(* Logix 5000 project; controller NWGG 1756-L72 rev 35.12; software revision 35.00; part 5 of 19 *)
(* tags used below, declared in another part *)
   _101AUTO : ALIAS FOR B9[101].4;
   _101HAND : ALIAS FOR B9[101].3;
   _101M : ALIAS FOR O25[9].3;
   _101MB : ALIAS FOR B9[101].2;
   _101STB : ALIAS FOR B9[101].0;
   _101STPB : ALIAS FOR B9[101].1;
   _101Y : ALIAS FOR I25[1].3;
   _102AUTO : ALIAS FOR B9[102].4;
   _102HAND : ALIAS FOR B9[102].3;
   _102M : ALIAS FOR O25[8].9;
   _102MB : ALIAS FOR B9[102].2;
   _102STB : ALIAS FOR B9[102].0;
   _102STPB : ALIAS FOR B9[102].1;
   _102Y : ALIAS FOR I25[0].9;
   _103AUTO : ALIAS FOR B9[103].4;
   _103HAND : ALIAS FOR B9[103].3;
   _103M : ALIAS FOR O25[8].12;
   _103MB : ALIAS FOR B9[103].2;
   _103STB : ALIAS FOR B9[103].0;
   _103STPB : ALIAS FOR B9[103].1;
   _103Y : ALIAS FOR I25[0].12;
   _106AUTO : ALIAS FOR B9[106].4;
   _106HAND : ALIAS FOR B9[106].3;
   _106M : ALIAS FOR O25[9].5;
   _106MB : ALIAS FOR B9[106].2;
   _106Y : ALIAS FOR I25[1].5;
   _107AUTO : ALIAS FOR B9[107].4;
   _107HAND : ALIAS FOR B9[107].3;
   _107M : ALIAS FOR O25[9].12;
   _107MB : ALIAS FOR B9[107].2;
   _107PS : ALIAS FOR I25[4].2;
   _107PSB : ALIAS FOR B9[107].5;
   _107STB : ALIAS FOR B9[107].0;
   _107STPB : ALIAS FOR B9[107].1;
   _107Y : ALIAS FOR I25[1].12;
   _108AUTO : ALIAS FOR B9[108].4;
   _108HAND : ALIAS FOR B9[108].3;
   _108M : ALIAS FOR O25[10].15;
   _108MB : ALIAS FOR B9[108].2;
   _108PS : ALIAS FOR I25[4].1;
   _108STB : ALIAS FOR B9[108].0;
   _108STPB : ALIAS FOR B9[108].1;
   _108Y : ALIAS FOR I25[2].15;
   _109_PS_DLY : ALIAS FOR T11[4];
   _109_SLOW_D : ALIAS FOR T11[5];
   _109_SLW_SP : ALIAS FOR I25[3].14;
   _109_STOP_D : ALIAS FOR T11[6];
   _109_STP_SP : ALIAS FOR I25[3].15;
   _109AUTO : ALIAS FOR B9[109].4;
   _109HAND : ALIAS FOR B9[109].3;
   _109M : ALIAS FOR O25[10].9;
   _109MB : ALIAS FOR B9[109].2;
   _109PS : ALIAS FOR I25[4].0;
   _109STB : ALIAS FOR B9[109].0;
   _109STPB : ALIAS FOR B9[109].1;
   _109Y : ALIAS FOR I25[2].9;
   _110AUTO : ALIAS FOR B9[110].4;
   _110HAND : ALIAS FOR B9[110].3;
   _110M : ALIAS FOR O25[8].15;
   _110MB : ALIAS FOR B9[110].2;
   _110STB : ALIAS FOR B9[110].0;
   _110STPB : ALIAS FOR B9[110].1;
   _110Y : ALIAS FOR I25[0].15;
   _111AUTO : ALIAS FOR B9[111].4;
   _111HAND : ALIAS FOR B9[111].3;
   _111M : ALIAS FOR O25[9].0;
   _111MB : ALIAS FOR B9[111].2;
   _111STB : ALIAS FOR B9[111].0;
   _111STPB : ALIAS FOR B9[111].1;
   _111Y : ALIAS FOR I25[1].0;
   _113AUTO : ALIAS FOR B9[113].4;
   _113HAND : ALIAS FOR B9[113].3;
   _113M : ALIAS FOR O25[10].5;
   _113MB : ALIAS FOR B9[113].2;
   _113STB : ALIAS FOR B9[113].0;
   _113STPB : ALIAS FOR B9[113].1;
   _113Y : ALIAS FOR I25[2].5;
   _116AUTO : ALIAS FOR B9[116].4;
   _116HAND : ALIAS FOR B9[116].3;
   _116M : ALIAS FOR O25[10].10;
   _116MB : ALIAS FOR B9[116].2;
   _116STB : ALIAS FOR B9[116].0;
   _116STPB : ALIAS FOR B9[116].1;
   _116Y : ALIAS FOR I25[2].10;
   _117AUTO : ALIAS FOR B9[117].4;
   _117HAND : ALIAS FOR B9[117].3;
   _117M : ALIAS FOR O25[10].8;
   _117MB : ALIAS FOR B9[117].2;
   _117STB : ALIAS FOR B9[117].0;
   _117STPB : ALIAS FOR B9[117].1;
   _117Y : ALIAS FOR I25[2].8;
   _11_PS : ALIAS FOR I25[4].14;
   _11_PS_DLY : ALIAS FOR T11[2];
   _11_SLOW_SP : ALIAS FOR I25[4].3;
   _11_STOP_SP : ALIAS FOR I25[4].6;
   _11AUTO : ALIAS FOR B9[11].4;
   _11HAND : ALIAS FOR B9[11].3;
   _11M : ALIAS FOR O25[9].2;
   _11MB : ALIAS FOR B9[11].2;
   _11STB : ALIAS FOR B9[11].0;
   _11STPB : ALIAS FOR B9[11].1;
   _11Y : ALIAS FOR I25[1].2;
   _122AUTO : ALIAS FOR B9[122].4;
   _122HAND : ALIAS FOR B9[122].3;
   _122M : ALIAS FOR O25[9].1;
   _122MB : ALIAS FOR B9[122].2;
   _122STB : ALIAS FOR B9[122].0;
   _122STPB : ALIAS FOR B9[122].1;
   _122Y : ALIAS FOR I25[1].1;
   _123_COMPUW : ALIAS FOR I18[7];
   _123_COMPUW1 : ALIAS FOR N7[20];
   _123AUTO : ALIAS FOR B9[123].4;
   _123HAND : ALIAS FOR B9[123].3;
   _123M : ALIAS FOR O25[10].6;
   _123MB : ALIAS FOR B9[123].2;
   _123STB : ALIAS FOR B9[123].0;
   _123STPB : ALIAS FOR B9[123].1;
   _123Y : ALIAS FOR I25[2].6;
   _124M : ALIAS FOR O25[9].13;
   _1AUTO : ALIAS FOR B9[1].4;
   _1HAND : ALIAS FOR B9[1].3;
   _1M : ALIAS FOR O25[9].8;
   _1MB : ALIAS FOR B9[1].2;
   _1STB : ALIAS FOR B9[1].0;
   _1STPB : ALIAS FOR B9[1].1;
   _1Y : ALIAS FOR I25[1].8;
   _25_16_0 : ALIAS FOR N200[10];
   _25_16_1 : ALIAS FOR N200[11];
   _25_16_2 : ALIAS FOR N200[12];
   _25_16_3 : ALIAS FOR N200[13];
   _2AUTO : ALIAS FOR B9[2].4;
   _2HAND : ALIAS FOR B9[2].3;
   _2M : ALIAS FOR O25[9].15;
   _2MB : ALIAS FOR B9[2].2;
   _2STB : ALIAS FOR B9[2].0;
   _2STPB : ALIAS FOR B9[2].1;
   _2Y : ALIAS FOR I25[1].15;
   _35AUTO : ALIAS FOR B9[35].4;
   _35HAND : ALIAS FOR B9[35].3;
   _35M : ALIAS FOR O25[10].13;
   _35MB : ALIAS FOR B9[35].2;
   _35STB : ALIAS FOR B9[35].0;
   _35STPB : ALIAS FOR B9[35].1;
   _35Y : ALIAS FOR I25[2].13;
   _36_FREQ_IN : ALIAS FOR N7[1];
   _36_FREQ_OU : ALIAS FOR N7[3];
   _36_SET_SPD : ALIAS FOR N7[2];
   _36_VFD_TO : ALIAS FOR N180[0];
   _36M : ALIAS FOR O25[8].0;
   _36RAUTO : ALIAS FOR B9[36].4;
   _36RHAND : ALIAS FOR B9[36].3;
   _36RMB : ALIAS FOR B9[36].2;
   _36RSTB : ALIAS FOR B9[36].0;
   _36RSTPB : ALIAS FOR B9[36].1;
   _36Y : ALIAS FOR I25[0].0;
   _3AUTO : ALIAS FOR B9[3].4;
   _3HAND : ALIAS FOR B9[3].3;
   _3M : ALIAS FOR O25[10].0;
   _3MB : ALIAS FOR B9[3].2;
   _3STB : ALIAS FOR B9[3].0;
   _3STPB : ALIAS FOR B9[3].1;
   _3Y : ALIAS FOR I25[2].0;
   _42AUTO : ALIAS FOR B9[42].4;
   _42HAND : ALIAS FOR B9[42].3;
   _42M : ALIAS FOR O25[11].1;
   _42MB : ALIAS FOR B9[42].2;
   _42STB : ALIAS FOR B9[42].0;
   _42STPB : ALIAS FOR B9[42].1;
   _42Y : ALIAS FOR I25[3].1;
   _43_ACC_WEI : ALIAS FOR C5[1].ACC;
   _43_BINDICA : ALIAS FOR B9[43].5;
   _43_RESET_C : ALIAS FOR B9[43].6;
   _43_SCREEN : ALIAS FOR C5[1];
   _43_SCREENI : ALIAS FOR I7.14;
   _43_WEIGHT : ALIAS FOR N7[0];
   _43AUTO : ALIAS FOR B9[43].4;
   _43HAND : ALIAS FOR B9[43].3;
   _43M : ALIAS FOR O25[10].14;
   _43MB : ALIAS FOR B9[43].2;
   _43STB : ALIAS FOR B9[43].0;
   _43STPB : ALIAS FOR B9[43].1;
   _43Y : ALIAS FOR I25[2].14;
   _47AUTO : ALIAS FOR B9[47].4;
   _47HAND : ALIAS FOR B9[47].3;
   _47M : ALIAS FOR O25[9].10;
   _47MB : ALIAS FOR B9[47].2;
   _47STB : ALIAS FOR B9[47].0;
   _47STPB : ALIAS FOR B9[47].1;
   _47Y : ALIAS FOR I25[1].10;
   _48_FREQ_IN : ALIAS FOR N7[10];
   _48_FREQ_OU : ALIAS FOR N7[12];
   _48_SET_SPD : ALIAS FOR N7[11];
   _48_VFD_TO : ALIAS FOR N180[2];
   _48AUTO : ALIAS FOR B9[48].4;
   _48HAND : ALIAS FOR B9[48].3;
   _48M : ALIAS FOR O25[8].3;
   _48MB : ALIAS FOR B9[48].2;
   _48STB : ALIAS FOR B9[48].0;
   _48STPB : ALIAS FOR B9[48].1;
   _48Y : ALIAS FOR I25[0].3;
   _49AUTO : ALIAS FOR B9[49].4;
   _49HAND : ALIAS FOR B9[49].3;
   _49M : ALIAS FOR O25[9].9;
   _49MB : ALIAS FOR B9[49].2;
   _49STB : ALIAS FOR B9[49].0;
   _49STPB : ALIAS FOR B9[49].1;
   _49Y : ALIAS FOR I25[1].9;
   _4AUTO : ALIAS FOR B9[4].4;
   _4HAND : ALIAS FOR B9[4].3;
   _4M : ALIAS FOR O25[10].1;
   _4MB : ALIAS FOR B9[4].2;
   _4STB : ALIAS FOR B9[4].0;
   _4STPB : ALIAS FOR B9[4].1;
   _4Y : ALIAS FOR I25[2].1;
   _50AUTO : ALIAS FOR B9[50].4;
   _50HAND : ALIAS FOR B9[50].3;
   _50M : ALIAS FOR O25[8].14;
   _50MB : ALIAS FOR B9[50].2;
   _50STB : ALIAS FOR B9[50].0;
   _50STPB : ALIAS FOR B9[50].1;
   _50Y : ALIAS FOR I25[0].14;
   _51_FREQ_IN : ALIAS FOR N7[13];
   _51_FREQ_OU : ALIAS FOR N7[15];
   _51_SET_SPD : ALIAS FOR N7[14];
   _51_VFD_TO : ALIAS FOR N180[3];
   _51AUTO : ALIAS FOR B9[51].4;
   _51HAND : ALIAS FOR B9[51].3;
   _51M : ALIAS FOR O25[8].4;
   _51MB : ALIAS FOR B9[51].2;
   _51STB : ALIAS FOR B9[51].0;
   _51STPB : ALIAS FOR B9[51].1;
   _51Y : ALIAS FOR I25[0].4;
   _52_FREQ_IN : ALIAS FOR N7[16];
   _52_FREQ_OU : ALIAS FOR N7[18];
   _52_SET_SPD : ALIAS FOR N7[17];
   _52AUTO : ALIAS FOR B9[52].4;
   _52HAND : ALIAS FOR B9[52].3;
   _52M : ALIAS FOR O25[8].6;
   _52MB : ALIAS FOR B9[52].2;
   _52STB : ALIAS FOR B9[52].0;
   _52STPB : ALIAS FOR B9[52].1;
   _52Y : ALIAS FOR I25[0].6;
   _53_FREQ_IN : ALIAS FOR N7[7];
   _53_FREQ_OU : ALIAS FOR N7[9];
   _53_SET_SPD : ALIAS FOR N7[8];
   _53_VFD_TO : ALIAS FOR N180[1];
   _53AUTO : ALIAS FOR B9[53].4;
   _53HAND : ALIAS FOR B9[53].3;
   _53M : ALIAS FOR O25[8].2;
   _53MB : ALIAS FOR B9[53].2;
(* _2_MAIN, continued *)

ROUTINE _09_SEED_MTR_9   (* ladder *)
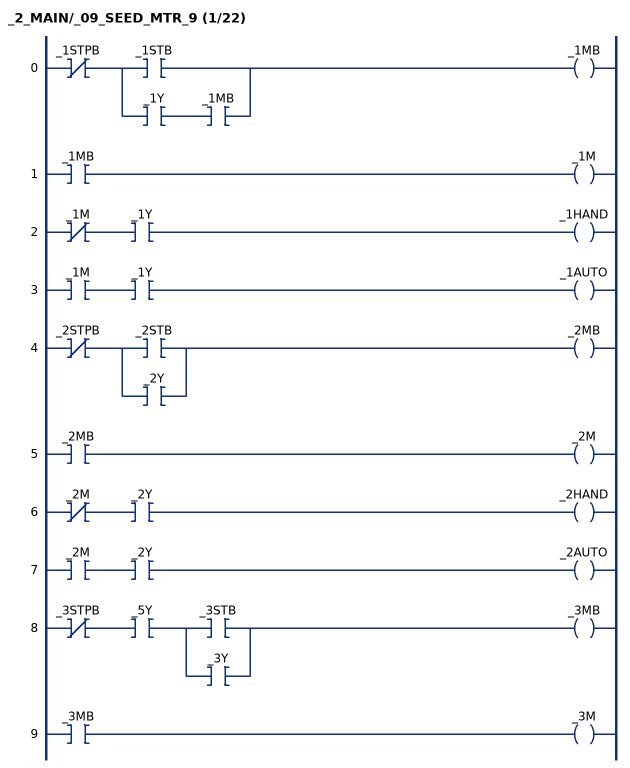
   0: XIO(_1STPB)[XIC(_1STB) ,XIC(_1Y) XIC(_1MB) ]OTE(_1MB);
   1: XIC(_1MB)OTE(_1M);
   2: XIO(_1M)XIC(_1Y)OTE(_1HAND);
   3: XIC(_1M)XIC(_1Y)OTE(_1AUTO);
   4: XIO(_2STPB)[XIC(_2STB) ,XIC(_2Y) ]OTE(_2MB);
   5: XIC(_2MB)OTE(_2M);
   6: XIO(_2M)XIC(_2Y)OTE(_2HAND);
   7: XIC(_2M)XIC(_2Y)OTE(_2AUTO);
   8: XIO(_3STPB)XIC(_5Y)[XIC(_3STB) ,XIC(_3Y) ]OTE(_3MB);
   9: XIC(_3MB)OTE(_3M);
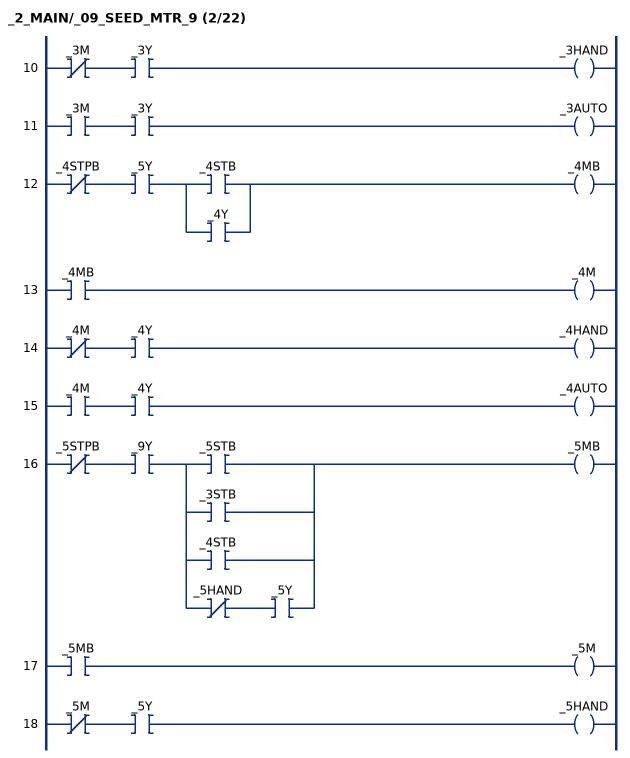
   10: XIO(_3M)XIC(_3Y)OTE(_3HAND);
   11: XIC(_3M)XIC(_3Y)OTE(_3AUTO);
   12: XIO(_4STPB)XIC(_5Y)[XIC(_4STB) ,XIC(_4Y) ]OTE(_4MB);
   13: XIC(_4MB)OTE(_4M);
   14: XIO(_4M)XIC(_4Y)OTE(_4HAND);
   15: XIC(_4M)XIC(_4Y)OTE(_4AUTO);
   16: XIO(_5STPB)XIC(_9Y)[XIC(_5STB) ,XIC(_3STB) ,XIC(_4STB) ,XIO(_5HAND) XIC(_5Y) ]OTE(_5MB);
   17: XIC(_5MB)OTE(_5M);
   18: XIO(_5M)XIC(_5Y)OTE(_5HAND);
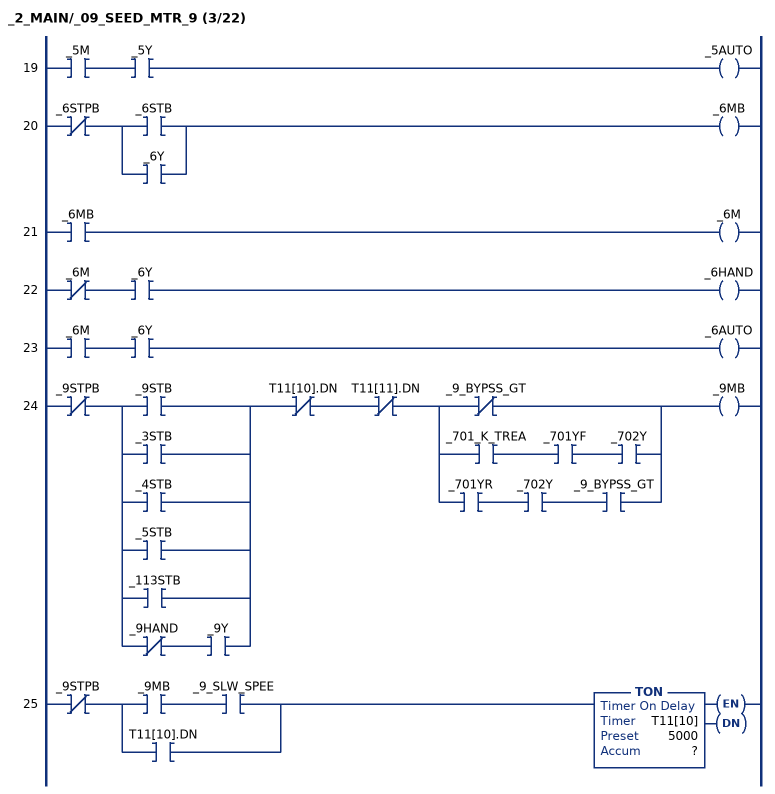
   19: XIC(_5M)XIC(_5Y)OTE(_5AUTO);
   20: XIO(_6STPB)[XIC(_6STB) ,XIC(_6Y) ]OTE(_6MB);
   21: XIC(_6MB)OTE(_6M);
   22: XIO(_6M)XIC(_6Y)OTE(_6HAND);
   23: XIC(_6M)XIC(_6Y)OTE(_6AUTO);
   24: XIO(_9STPB)[XIC(_9STB) ,XIC(_3STB) ,XIC(_4STB) ,XIC(_5STB) ,XIC(_113STB) ,XIO(_9HAND) XIC(_9Y) ]XIO(T11[10].DN)XIO(T11[11].DN)[XIO(_9_BYPSS_GT) ,XIC(_701_K_TREA) XIC(_701YF) XIC(_702Y) ,XIC(_701YR) XIC(_702Y) XIC(_9_BYPSS_GT) ]OTE(_9MB);
   25: XIO(_9STPB)[XIC(_9MB) XIC(_9_SLW_SPEE) ,XIC(T11[10].DN) ]TON(T11[10],?,?);
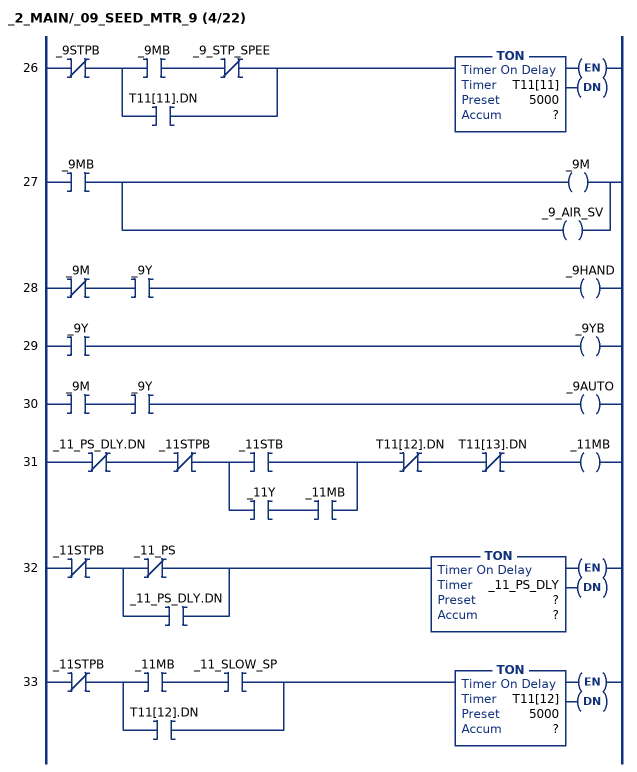
   26: XIO(_9STPB)[XIC(_9MB) XIO(_9_STP_SPEE) ,XIC(T11[11].DN) ]TON(T11[11],?,?);
   27: XIC(_9MB)[OTE(_9M) ,OTE(_9_AIR_SV) ];
   28: XIO(_9M)XIC(_9Y)OTE(_9HAND);
   29: XIC(_9Y)OTE(_9YB);
   30: XIC(_9M)XIC(_9Y)OTE(_9AUTO);
   31: XIO(_11_PS_DLY.DN)XIO(_11STPB)[XIC(_11STB) ,XIC(_11Y) XIC(_11MB) ]XIO(T11[12].DN)XIO(T11[13].DN)OTE(_11MB);
   32: XIO(_11STPB)[XIO(_11_PS) ,XIC(_11_PS_DLY.DN) ]TON(_11_PS_DLY,?,?);
   33: XIO(_11STPB)[XIC(_11MB) XIC(_11_SLOW_SP) ,XIC(T11[12].DN) ]TON(T11[12],?,?);
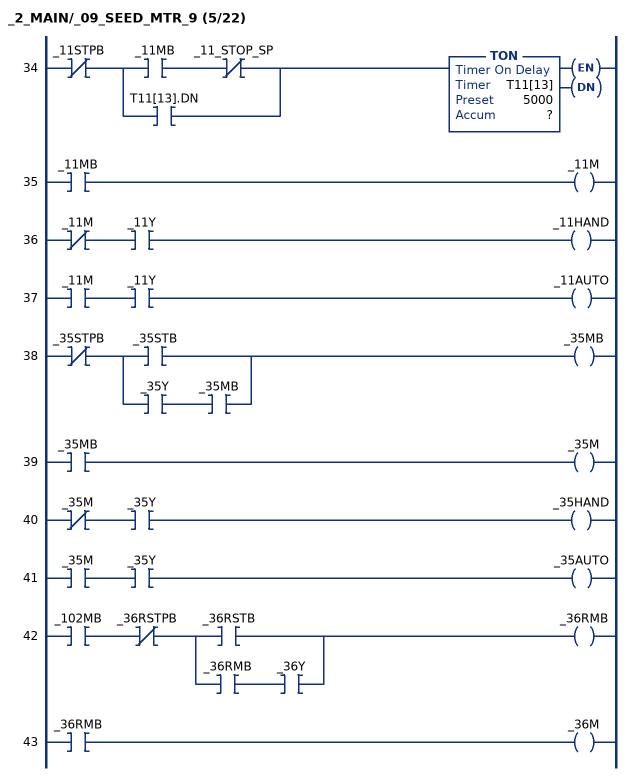
   34: XIO(_11STPB)[XIC(_11MB) XIO(_11_STOP_SP) ,XIC(T11[13].DN) ]TON(T11[13],?,?);
   35: XIC(_11MB)OTE(_11M);
   36: XIO(_11M)XIC(_11Y)OTE(_11HAND);
   37: XIC(_11M)XIC(_11Y)OTE(_11AUTO);
   38: XIO(_35STPB)[XIC(_35STB) ,XIC(_35Y) XIC(_35MB) ]OTE(_35MB);
   39: XIC(_35MB)OTE(_35M);
   40: XIO(_35M)XIC(_35Y)OTE(_35HAND);
   41: XIC(_35M)XIC(_35Y)OTE(_35AUTO);
   42: XIC(_102MB)XIO(_36RSTPB)[XIC(_36RSTB) ,XIC(_36RMB) XIC(_36Y) ]OTE(_36RMB);
   43: XIC(_36RMB)OTE(_36M);
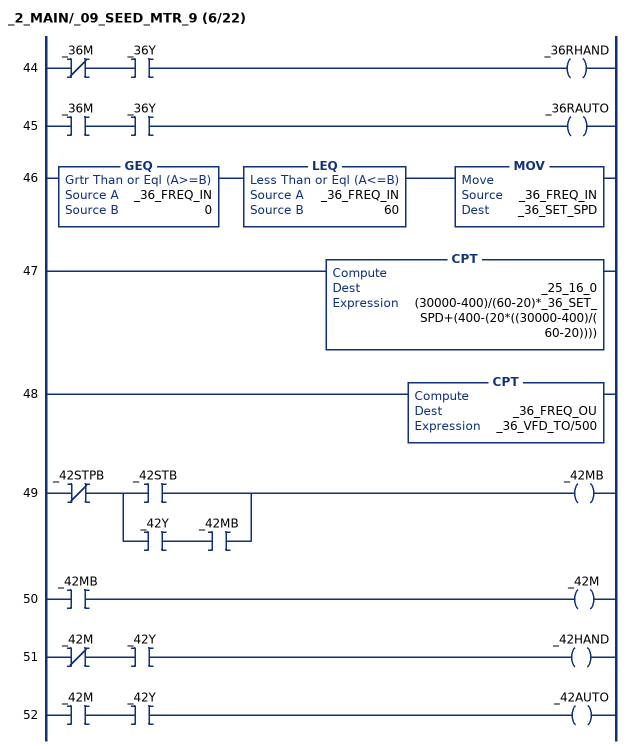
   44: XIO(_36M)XIC(_36Y)OTE(_36RHAND);
   45: XIC(_36M)XIC(_36Y)OTE(_36RAUTO);
   46: GEQ(_36_FREQ_IN,0)LEQ(_36_FREQ_IN,60)MOV(_36_FREQ_IN,_36_SET_SPD);
   47: CPT(_25_16_0,(30000-400)/(60-20)*_36_SET_SPD+(400-(20*((30000-400)/(60-20)))));
   48: CPT(_36_FREQ_OU,_36_VFD_TO/500);
   49: XIO(_42STPB)[XIC(_42STB) ,XIC(_42Y) XIC(_42MB) ]OTE(_42MB);
   50: XIC(_42MB)OTE(_42M);
   51: XIO(_42M)XIC(_42Y)OTE(_42HAND);
   52: XIC(_42M)XIC(_42Y)OTE(_42AUTO);
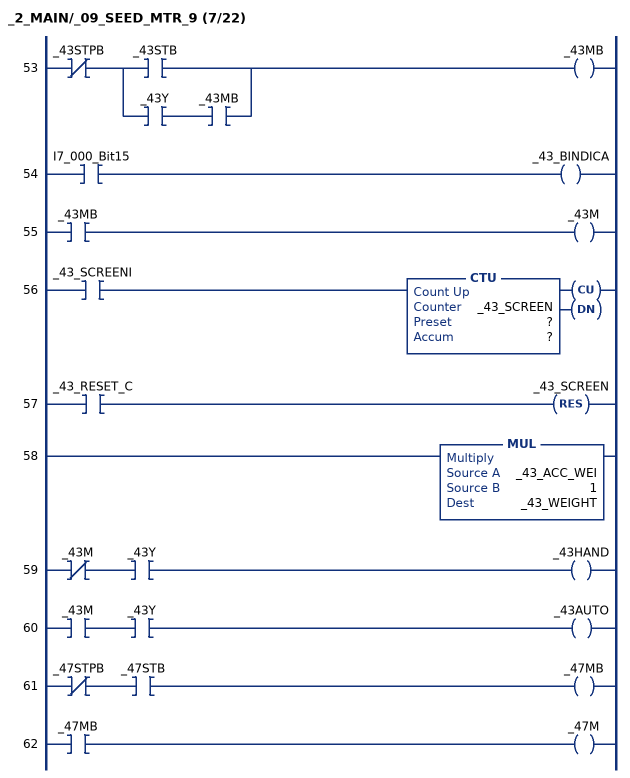
   53: XIO(_43STPB)[XIC(_43STB) ,XIC(_43Y) XIC(_43MB) ]OTE(_43MB);
   54: XIC(I7_000_Bit15)OTE(_43_BINDICA);
   55: XIC(_43MB)OTE(_43M);
   56: XIC(_43_SCREENI)CTU(_43_SCREEN,?,?);
   57: XIC(_43_RESET_C)RES(_43_SCREEN);
   58: MUL(_43_ACC_WEI,1,_43_WEIGHT);
   59: XIO(_43M)XIC(_43Y)OTE(_43HAND);
   60: XIC(_43M)XIC(_43Y)OTE(_43AUTO);
   61: XIO(_47STPB)XIC(_47STB)OTE(_47MB);
   62: XIC(_47MB)OTE(_47M);
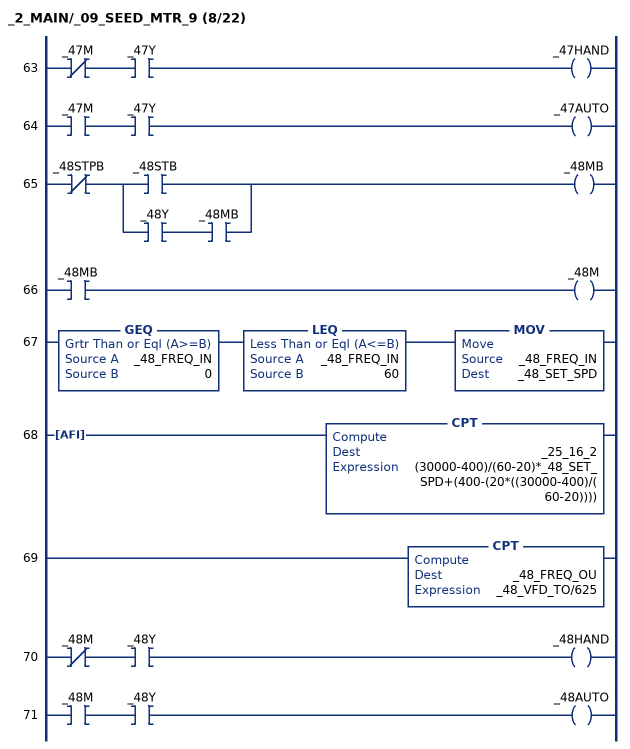
   63: XIO(_47M)XIC(_47Y)OTE(_47HAND);
   64: XIC(_47M)XIC(_47Y)OTE(_47AUTO);
   65: XIO(_48STPB)[XIC(_48STB) ,XIC(_48Y) XIC(_48MB) ]OTE(_48MB);
   66: XIC(_48MB)OTE(_48M);
   67: GEQ(_48_FREQ_IN,0)LEQ(_48_FREQ_IN,60)MOV(_48_FREQ_IN,_48_SET_SPD);
   68: AFI()CPT(_25_16_2,(30000-400)/(60-20)*_48_SET_SPD+(400-(20*((30000-400)/(60-20)))));
   69: CPT(_48_FREQ_OU,_48_VFD_TO/625);
   70: XIO(_48M)XIC(_48Y)OTE(_48HAND);
   71: XIC(_48M)XIC(_48Y)OTE(_48AUTO);
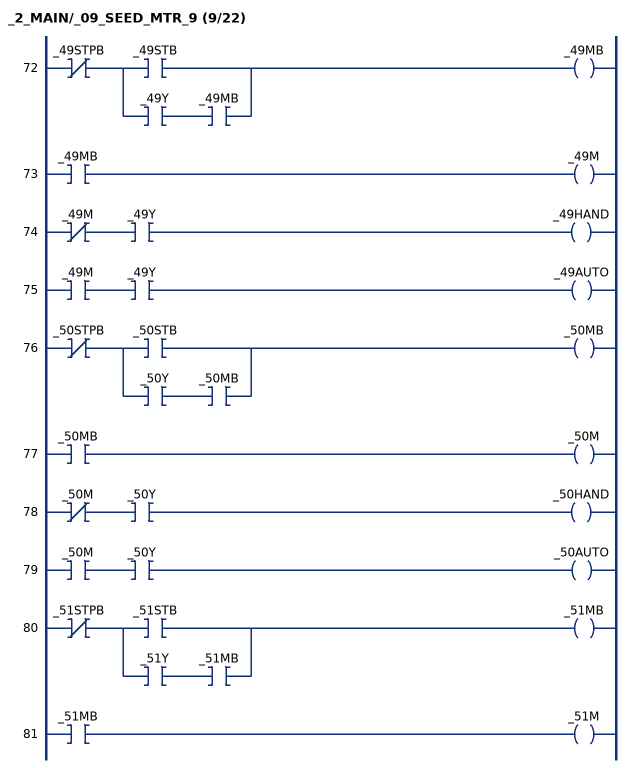
   72: XIO(_49STPB)[XIC(_49STB) ,XIC(_49Y) XIC(_49MB) ]OTE(_49MB);
   73: XIC(_49MB)OTE(_49M);
   74: XIO(_49M)XIC(_49Y)OTE(_49HAND);
   75: XIC(_49M)XIC(_49Y)OTE(_49AUTO);
   76: XIO(_50STPB)[XIC(_50STB) ,XIC(_50Y) XIC(_50MB) ]OTE(_50MB);
   77: XIC(_50MB)OTE(_50M);
   78: XIO(_50M)XIC(_50Y)OTE(_50HAND);
   79: XIC(_50M)XIC(_50Y)OTE(_50AUTO);
   80: XIO(_51STPB)[XIC(_51STB) ,XIC(_51Y) XIC(_51MB) ]OTE(_51MB);
   81: XIC(_51MB)OTE(_51M);
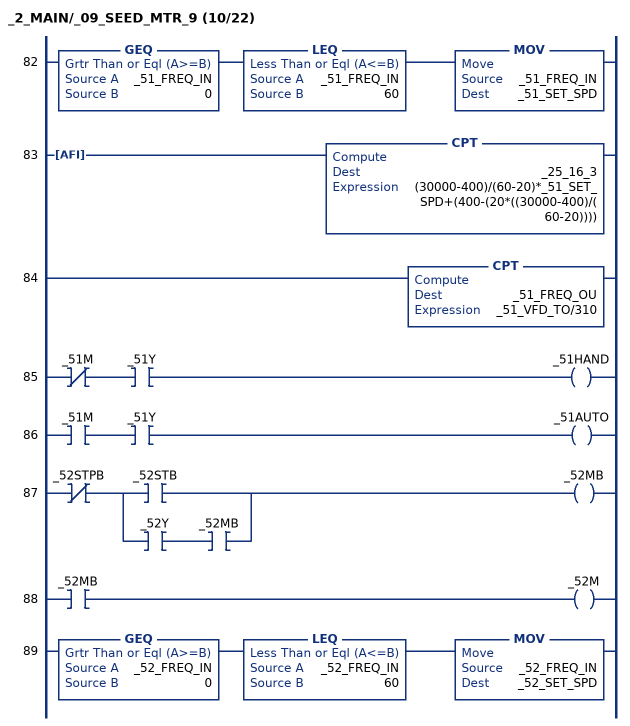
   82: GEQ(_51_FREQ_IN,0)LEQ(_51_FREQ_IN,60)MOV(_51_FREQ_IN,_51_SET_SPD);
   83: AFI()CPT(_25_16_3,(30000-400)/(60-20)*_51_SET_SPD+(400-(20*((30000-400)/(60-20)))));
   84: CPT(_51_FREQ_OU,_51_VFD_TO/310);
   85: XIO(_51M)XIC(_51Y)OTE(_51HAND);
   86: XIC(_51M)XIC(_51Y)OTE(_51AUTO);
   87: XIO(_52STPB)[XIC(_52STB) ,XIC(_52Y) XIC(_52MB) ]OTE(_52MB);
   88: XIC(_52MB)OTE(_52M);
   89: GEQ(_52_FREQ_IN,0)LEQ(_52_FREQ_IN,60)MOV(_52_FREQ_IN,_52_SET_SPD);
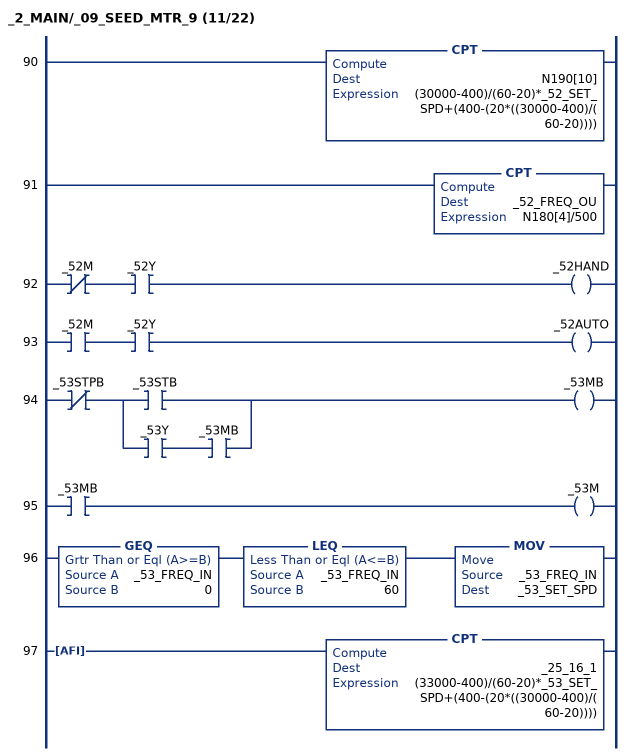
   90: CPT(N190[10],(30000-400)/(60-20)*_52_SET_SPD+(400-(20*((30000-400)/(60-20)))));
   91: CPT(_52_FREQ_OU,N180[4]/500);
   92: XIO(_52M)XIC(_52Y)OTE(_52HAND);
   93: XIC(_52M)XIC(_52Y)OTE(_52AUTO);
   94: XIO(_53STPB)[XIC(_53STB) ,XIC(_53Y) XIC(_53MB) ]OTE(_53MB);
   95: XIC(_53MB)OTE(_53M);
   96: GEQ(_53_FREQ_IN,0)LEQ(_53_FREQ_IN,60)MOV(_53_FREQ_IN,_53_SET_SPD);
   97: AFI()CPT(_25_16_1,(33000-400)/(60-20)*_53_SET_SPD+(400-(20*((30000-400)/(60-20)))));
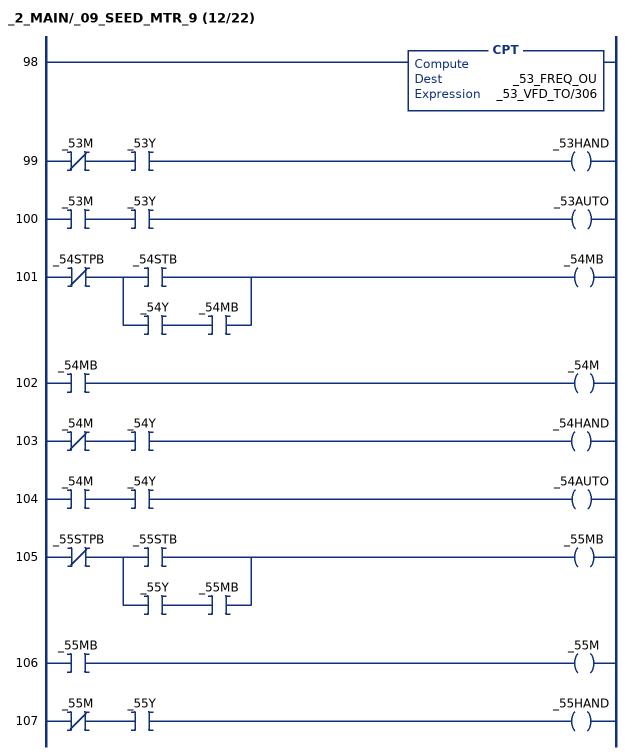
   98: CPT(_53_FREQ_OU,_53_VFD_TO/306);
   99: XIO(_53M)XIC(_53Y)OTE(_53HAND);
   100: XIC(_53M)XIC(_53Y)OTE(_53AUTO);
   101: XIO(_54STPB)[XIC(_54STB) ,XIC(_54Y) XIC(_54MB) ]OTE(_54MB);
   102: XIC(_54MB)OTE(_54M);
   103: XIO(_54M)XIC(_54Y)OTE(_54HAND);
   104: XIC(_54M)XIC(_54Y)OTE(_54AUTO);
   105: XIO(_55STPB)[XIC(_55STB) ,XIC(_55Y) XIC(_55MB) ]OTE(_55MB);
   106: XIC(_55MB)OTE(_55M);
   107: XIO(_55M)XIC(_55Y)OTE(_55HAND);
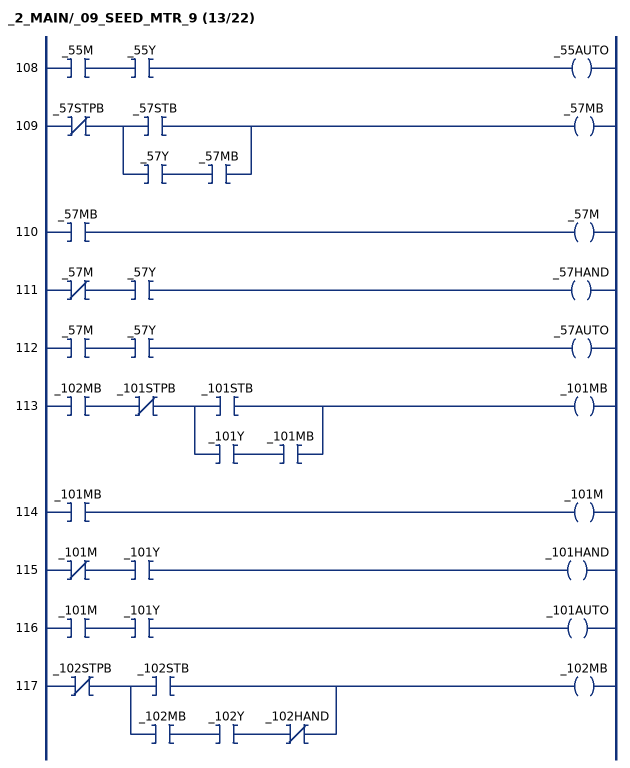
   108: XIC(_55M)XIC(_55Y)OTE(_55AUTO);
   109: XIO(_57STPB)[XIC(_57STB) ,XIC(_57Y) XIC(_57MB) ]OTE(_57MB);
   110: XIC(_57MB)OTE(_57M);
   111: XIO(_57M)XIC(_57Y)OTE(_57HAND);
   112: XIC(_57M)XIC(_57Y)OTE(_57AUTO);
   113: XIC(_102MB)XIO(_101STPB)[XIC(_101STB) ,XIC(_101Y) XIC(_101MB) ]OTE(_101MB);
   114: XIC(_101MB)OTE(_101M);
   115: XIO(_101M)XIC(_101Y)OTE(_101HAND);
   116: XIC(_101M)XIC(_101Y)OTE(_101AUTO);
   117: XIO(_102STPB)[XIC(_102STB) ,XIC(_102MB) XIC(_102Y) XIO(_102HAND) ]OTE(_102MB);
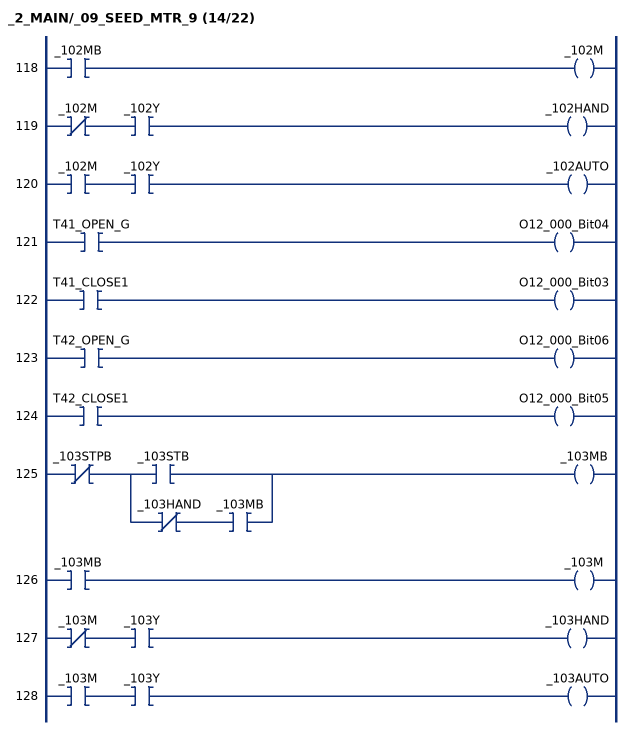
   118: XIC(_102MB)OTE(_102M);
   119: XIO(_102M)XIC(_102Y)OTE(_102HAND);
   120: XIC(_102M)XIC(_102Y)OTE(_102AUTO);
   121: XIC(T41_OPEN_G)OTE(O12_000_Bit04);
   122: XIC(T41_CLOSE1)OTE(O12_000_Bit03);
   123: XIC(T42_OPEN_G)OTE(O12_000_Bit06);
   124: XIC(T42_CLOSE1)OTE(O12_000_Bit05);
   125: XIO(_103STPB)[XIC(_103STB) ,XIO(_103HAND) XIC(_103MB) ]OTE(_103MB);
   126: XIC(_103MB)OTE(_103M);
   127: XIO(_103M)XIC(_103Y)OTE(_103HAND);
   128: XIC(_103M)XIC(_103Y)OTE(_103AUTO);
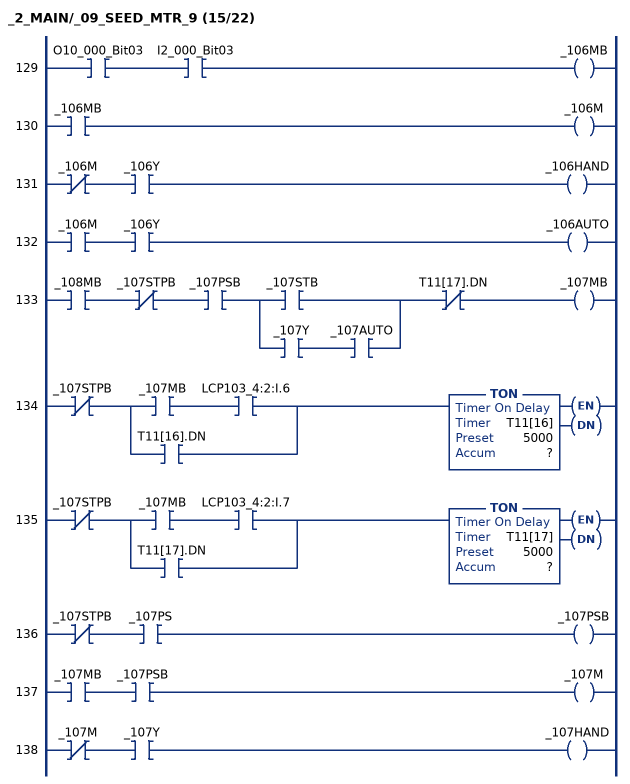
   129: XIC(O10_000_Bit03)XIC(I2_000_Bit03)OTE(_106MB);
   130: XIC(_106MB)OTE(_106M);
   131: XIO(_106M)XIC(_106Y)OTE(_106HAND);
   132: XIC(_106M)XIC(_106Y)OTE(_106AUTO);
   133: XIC(_108MB)XIO(_107STPB)XIC(_107PSB)[XIC(_107STB) ,XIC(_107Y) XIC(_107AUTO) ]XIO(T11[17].DN)OTE(_107MB);
   134: XIO(_107STPB)[XIC(_107MB) XIC(LCP103_4:2:I.6) ,XIC(T11[16].DN) ]TON(T11[16],?,?);
   135: XIO(_107STPB)[XIC(_107MB) XIC(LCP103_4:2:I.7) ,XIC(T11[17].DN) ]TON(T11[17],?,?);
   136: XIO(_107STPB)XIC(_107PS)OTE(_107PSB);
   137: XIC(_107MB)XIC(_107PSB)OTE(_107M);
   138: XIO(_107M)XIC(_107Y)OTE(_107HAND);
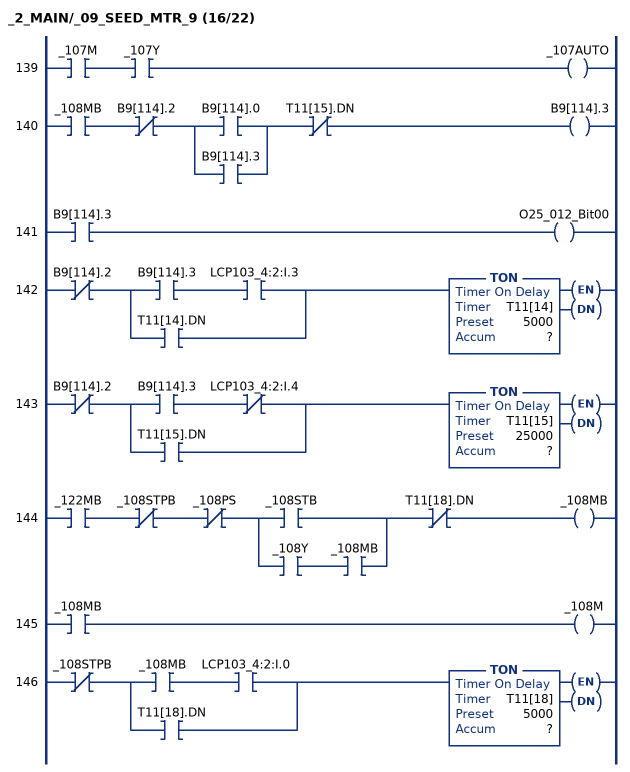
   139: XIC(_107M)XIC(_107Y)OTE(_107AUTO);
   140: XIC(_108MB)XIO(B9[114].2)[XIC(B9[114].0) ,XIC(B9[114].3) ]XIO(T11[15].DN)OTE(B9[114].3);
   141: XIC(B9[114].3)OTE(O25_012_Bit00);
   142: XIO(B9[114].2)[XIC(B9[114].3) XIC(LCP103_4:2:I.3) ,XIC(T11[14].DN) ]TON(T11[14],?,?);
   143: XIO(B9[114].2)[XIC(B9[114].3) XIO(LCP103_4:2:I.4) ,XIC(T11[15].DN) ]TON(T11[15],?,?);
   144: XIC(_122MB)XIO(_108STPB)XIO(_108PS)[XIC(_108STB) ,XIC(_108Y) XIC(_108MB) ]XIO(T11[18].DN)OTE(_108MB);
   145: XIC(_108MB)OTE(_108M);
   146: XIO(_108STPB)[XIC(_108MB) XIC(LCP103_4:2:I.0) ,XIC(T11[18].DN) ]TON(T11[18],?,?);
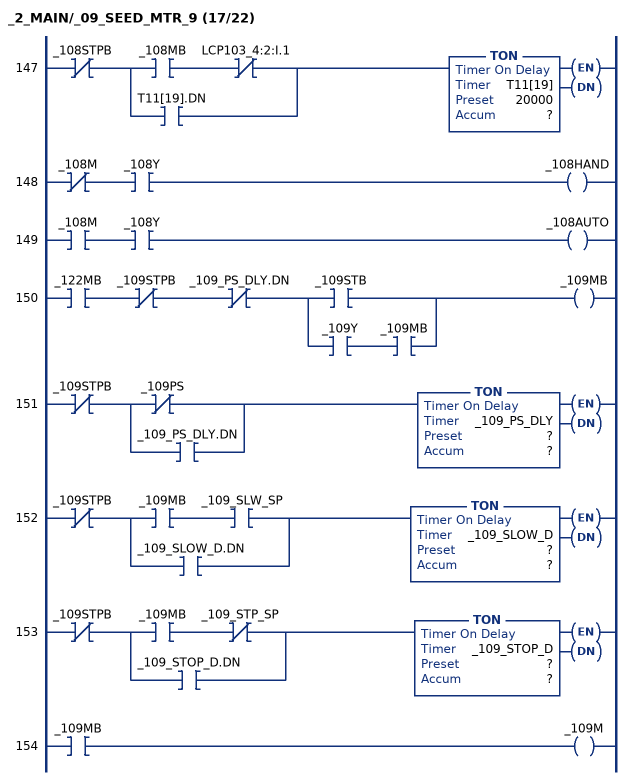
   147: XIO(_108STPB)[XIC(_108MB) XIO(LCP103_4:2:I.1) ,XIC(T11[19].DN) ]TON(T11[19],?,?);
   148: XIO(_108M)XIC(_108Y)OTE(_108HAND);
   149: XIC(_108M)XIC(_108Y)OTE(_108AUTO);
   150: XIC(_122MB)XIO(_109STPB)XIO(_109_PS_DLY.DN)[XIC(_109STB) ,XIC(_109Y) XIC(_109MB) ]OTE(_109MB);
   151: XIO(_109STPB)[XIO(_109PS) ,XIC(_109_PS_DLY.DN) ]TON(_109_PS_DLY,?,?);
   152: XIO(_109STPB)[XIC(_109MB) XIC(_109_SLW_SP) ,XIC(_109_SLOW_D.DN) ]TON(_109_SLOW_D,?,?);
   153: XIO(_109STPB)[XIC(_109MB) XIO(_109_STP_SP) ,XIC(_109_STOP_D.DN) ]TON(_109_STOP_D,?,?);
   154: XIC(_109MB)OTE(_109M);
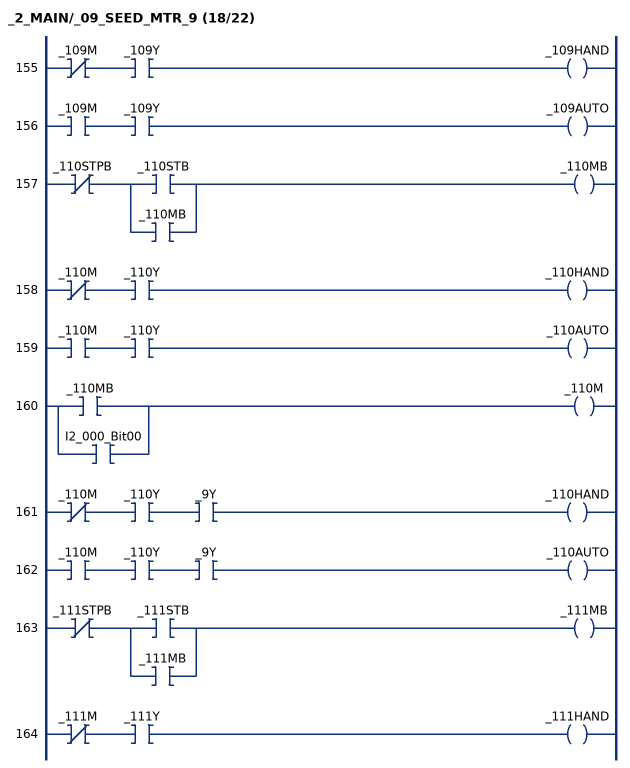
   155: XIO(_109M)XIC(_109Y)OTE(_109HAND);
   156: XIC(_109M)XIC(_109Y)OTE(_109AUTO);
   157: XIO(_110STPB)[XIC(_110STB) ,XIC(_110MB) ]OTE(_110MB);
   158: XIO(_110M)XIC(_110Y)OTE(_110HAND);
   159: XIC(_110M)XIC(_110Y)OTE(_110AUTO);
   160: [XIC(_110MB) ,XIC(I2_000_Bit00) ]OTE(_110M);
   161: XIO(_110M)XIC(_110Y)XIC(_9Y)OTE(_110HAND);
   162: XIC(_110M)XIC(_110Y)XIC(_9Y)OTE(_110AUTO);
   163: XIO(_111STPB)[XIC(_111STB) ,XIC(_111MB) ]OTE(_111MB);
   164: XIO(_111M)XIC(_111Y)OTE(_111HAND);
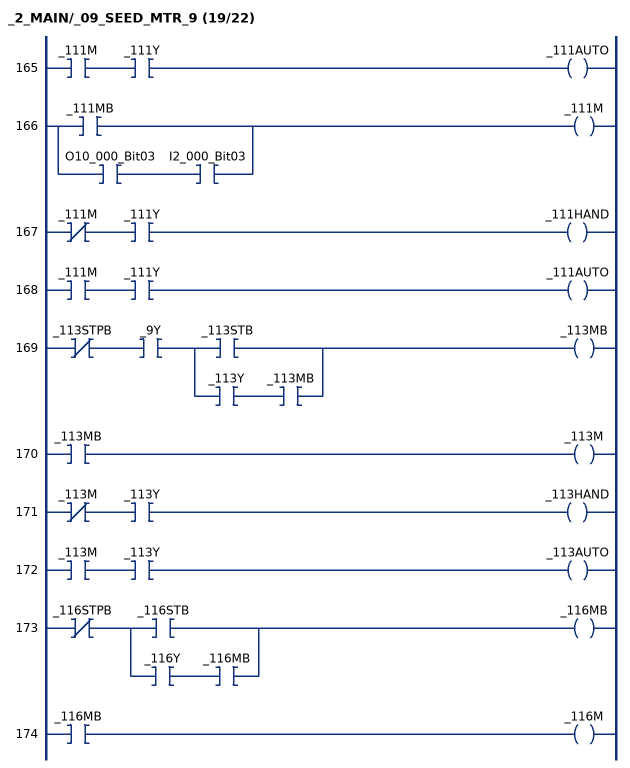
   165: XIC(_111M)XIC(_111Y)OTE(_111AUTO);
   166: [XIC(_111MB) ,XIC(O10_000_Bit03) XIC(I2_000_Bit03) ]OTE(_111M);
   167: XIO(_111M)XIC(_111Y)OTE(_111HAND);
   168: XIC(_111M)XIC(_111Y)OTE(_111AUTO);
   169: XIO(_113STPB)XIC(_9Y)[XIC(_113STB) ,XIC(_113Y) XIC(_113MB) ]OTE(_113MB);
   170: XIC(_113MB)OTE(_113M);
   171: XIO(_113M)XIC(_113Y)OTE(_113HAND);
   172: XIC(_113M)XIC(_113Y)OTE(_113AUTO);
   173: XIO(_116STPB)[XIC(_116STB) ,XIC(_116Y) XIC(_116MB) ]OTE(_116MB);
   174: XIC(_116MB)OTE(_116M);
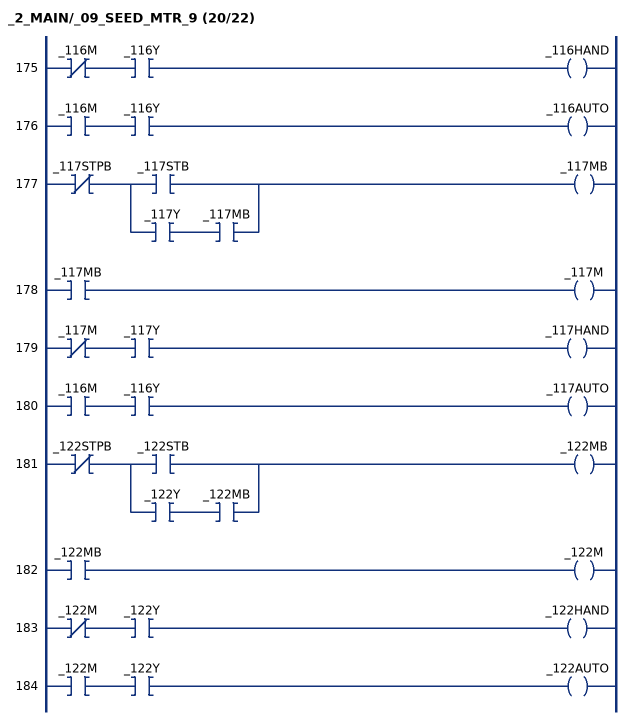
   175: XIO(_116M)XIC(_116Y)OTE(_116HAND);
   176: XIC(_116M)XIC(_116Y)OTE(_116AUTO);
   177: XIO(_117STPB)[XIC(_117STB) ,XIC(_117Y) XIC(_117MB) ]OTE(_117MB);
   178: XIC(_117MB)OTE(_117M);
   179: XIO(_117M)XIC(_117Y)OTE(_117HAND);
   180: XIC(_116M)XIC(_116Y)OTE(_117AUTO);
   181: XIO(_122STPB)[XIC(_122STB) ,XIC(_122Y) XIC(_122MB) ]OTE(_122MB);
   182: XIC(_122MB)OTE(_122M);
   183: XIO(_122M)XIC(_122Y)OTE(_122HAND);
   184: XIC(_122M)XIC(_122Y)OTE(_122AUTO);
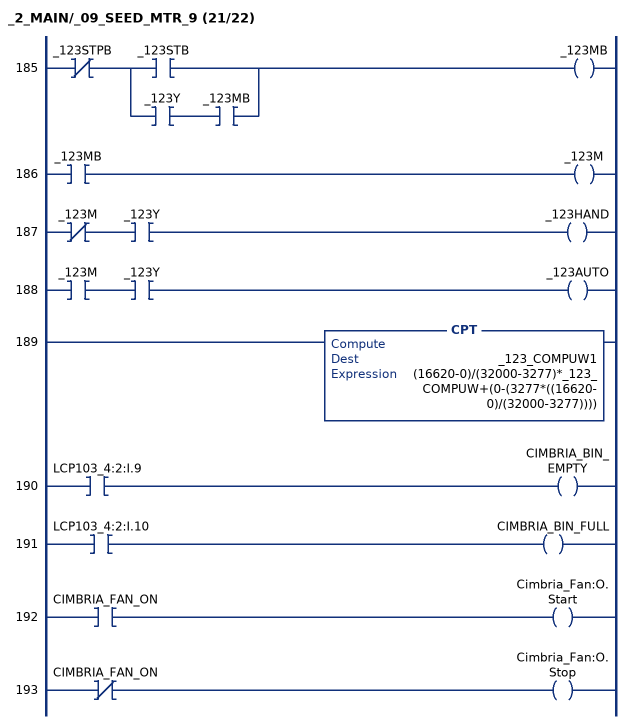
   185: XIO(_123STPB)[XIC(_123STB) ,XIC(_123Y) XIC(_123MB) ]OTE(_123MB);
   186: XIC(_123MB)OTE(_123M);
   187: XIO(_123M)XIC(_123Y)OTE(_123HAND);
   188: XIC(_123M)XIC(_123Y)OTE(_123AUTO);
   189: CPT(_123_COMPUW1,(16620-0)/(32000-3277)*_123_COMPUW+(0-(3277*((16620-0)/(32000-3277)))));
   190: XIC(LCP103_4:2:I.9)OTE(CIMBRIA_BIN_EMPTY);
   191: XIC(LCP103_4:2:I.10)OTE(CIMBRIA_BIN_FULL);
   192: XIC(CIMBRIA_FAN_ON)OTE(Cimbria_Fan:O.Start);
   193: XIO(CIMBRIA_FAN_ON)OTE(Cimbria_Fan:O.Stop);
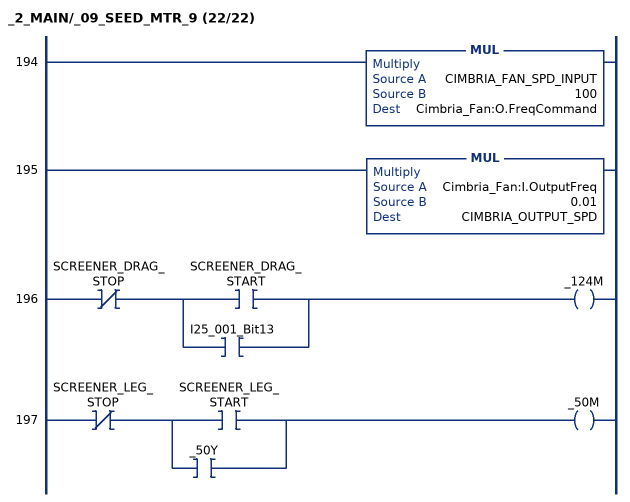
   194: MUL(CIMBRIA_FAN_SPD_INPUT,100,Cimbria_Fan:O.FreqCommand);
   195: MUL(Cimbria_Fan:I.OutputFreq,0.01,CIMBRIA_OUTPUT_SPD);
   196: XIO(SCREENER_DRAG_STOP)[XIC(SCREENER_DRAG_START) ,XIC(I25_001_Bit13) ]OTE(_124M);
   197: XIO(SCREENER_LEG_STOP)[XIC(SCREENER_LEG_START) ,XIC(_50Y) ]OTE(_50M);
END_ROUTINE
